(* PLC project AgentPLC, Beckhoff Automation GmbH TwinCAT PLC Control 3.5.21.61 *)
(* stored: creationDateTime 2026-11-03T09:46:44.5907528, modificationDateTime 2026-11-03T09:46:44.5943573 *)

PROGRAM MAIN
VAR
	Start : BOOL; // Offline test input
	Lamp : BOOL; // Offline test output
END_VAR

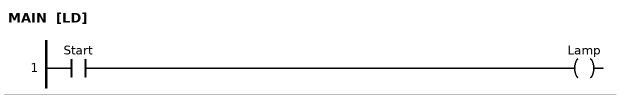
(* LD diagram, written out as Structured Text *)
(* Agent-authored native LD probe *)

Lamp := Start;
END_PROGRAM

CONFIGURATION Application
  RESOURCE AgentPLC ON PLC
    TASK PlcTask(INTERVAL := T#0ms, PRIORITY := 20);
    PROGRAM MAIN WITH PlcTask : MAIN;
  END_RESOURCE
END_CONFIGURATION
